FUNCTION_BLOCK "FB_UDP_Pasarela"
{ S7_Optimized_Access := 'TRUE' }
VERSION : 0.1
// PLC_Camara: 279 bloques (un Serialize por miembro de DB o tag). Generado por generar.py
   VAR_INPUT
      Deshabilitar : Bool := FALSE;
      Periodo : Time := T#100ms;
      Ip_pasarela : Array[1..4] of Byte := [172, 21, 0, 200];
      Puerto : UInt := 5000;
   END_VAR
   VAR_OUTPUT
      Conectado : Bool;
      Enviados : UDInt;
      Fallidos : UDInt;
      Bloques_omitidos : Int;
      Estado_tusend : Word;
      Estado_tcon : Word;
      Ultimo_error_tcon : Word;
      Errores_tcon : UDInt;
      Intentos_tcon : UDInt;
      Conexiones_ok : UDInt;
   END_VAR
   VAR
      Etapa : Int;
      Secuencia : UDInt;
      Marca_tiempo : LInt;
      Lanza_conexion : Bool;
      Flanco_conexion : R_TRIG;
      Lanza_envio : Bool;
      Conexion : TCON_IP_v4;
      Destino : TADDR_Param;
      Cliente_con : TCON;
      Cliente_envio : TUSEND;
      Espera_conexion : TON_TIME;
      Espera_periodo : TON_TIME;
      Espera_envio : TON_TIME;
      Datagrama : Array[0..1499] of Byte;
      Foto : Array[0..3384] of Byte;
      Total : DInt;
      Cursor : DInt;
      Bytes_trozo : DInt;
      Bloques_trozo : UInt;
      Bloques_escritos : Int;
      Copia_1 : Array[0..107] of Byte;
      Copia_2 : Bool;
      Copia_3 : Bool;
      Copia_4 : Bool;
      Copia_5 : Bool;
      Copia_6 : Bool;
      Copia_7 : Bool;
      Copia_8 : Bool;
      Copia_9 : Bool;
      Copia_10 : UDInt;
      Copia_11 : UDInt;
      Copia_12 : Bool;
      Copia_13 : Array[0..107] of Byte;
      Copia_14 : UDInt;
      Copia_15 : UDInt;
      Copia_16 : DWord;
      Copia_17 : DWord;
      Copia_18 : DWord;
      Copia_19 : DWord;
      Copia_20 : DWord;
      Copia_21 : DWord;
      Copia_22 : DWord;
      Copia_23 : DWord;
      Copia_24 : DWord;
      Copia_25 : DWord;
      Copia_26 : DWord;
      Copia_27 : DWord;
      Copia_28 : DWord;
      Copia_29 : DWord;
      Copia_30 : DWord;
      Copia_31 : DWord;
      Copia_32 : DWord;
      Copia_33 : DWord;
      Copia_34 : DWord;
      Copia_35 : DWord;
      Copia_36 : DWord;
      Copia_37 : DWord;
      Copia_38 : DWord;
      Copia_39 : DWord;
      Copia_40 : DWord;
      Copia_41 : DWord;
      Copia_42 : DWord;
      Copia_43 : DWord;
      Copia_44 : DWord;
      Copia_45 : DWord;
      Copia_46 : DWord;
      Copia_47 : DWord;
      Copia_48 : Bool;
      Copia_49 : DInt;
      Copia_50 : DInt;
      Copia_51 : Time;
      Copia_52 : "UDT_Entradas_Basico";
      Copia_53 : "UDT_Entradas_RFID";
      Copia_54 : "UDT_Entradas_Stopper";
      Copia_55 : Word;
      Copia_56 : Word;
      Copia_57 : Bool;
      Copia_58 : Bool;
      Copia_59 : Bool;
      Copia_60 : Bool;
      Copia_61 : Bool;
      Copia_62 : DWord;
      Copia_63 : DWord;
      Copia_64 : DWord;
      Copia_65 : DWord;
      Copia_66 : DWord;
      Copia_67 : DWord;
      Copia_68 : DWord;
      Copia_69 : DWord;
      Copia_70 : USInt;
      Copia_71 : UInt;
      Copia_72 : Bool;
      Copia_73 : DInt;
      Copia_74 : Bool;
      Copia_75 : Bool;
      Copia_76 : Bool;
      Copia_77 : UDInt;
      Copia_78 : UDInt;
      Copia_79 : DInt;
      Copia_80 : Int;
      Copia_81 : Bool;
      Copia_82 : Bool;
      Copia_83 : Bool;
      Copia_84 : Bool;
      Copia_85 : Bool;
      Copia_86 : Bool;
      Copia_87 : "UDT_Estado";
      Copia_88 : Bool;
      Copia_89 : Bool;
      Copia_90 : Bool;
      Copia_91 : Bool;
      Copia_92 : Bool;
      Copia_93 : Bool;
      Copia_94 : Bool;
      Copia_95 : Bool;
      Copia_96 : Bool;
      Copia_97 : Bool;
      Copia_98 : Int;
      Copia_99 : Int;
      Copia_100 : Int;
      Copia_101 : Bool;
      Copia_102 : Bool;
      Copia_103 : Bool;
      Copia_104 : Bool;
      Copia_105 : Bool;
      Copia_106 : Bool;
      Copia_107 : Bool;
      Copia_108 : Bool;
      Copia_109 : Bool;
      Copia_110 : Bool;
      Copia_111 : Bool;
      Copia_112 : Bool;
      Copia_113 : Bool;
      Copia_114 : Bool;
      Copia_115 : Bool;
      Copia_116 : Bool;
      Copia_117 : DInt;
      Copia_118 : DInt;
      Copia_119 : Bool;
      Copia_120 : Int;
      Copia_121 : Bool;
      Copia_122 : Bool;
      Copia_123 : Bool;
      Copia_124 : Bool;
      Copia_125 : Int;
      Copia_126 : Bool;
      Copia_127 : Bool;
      Copia_128 : Bool;
      Copia_129 : Bool;
      Copia_130 : Time;
      Copia_131 : Time;
      Copia_132 : Bool;
      Copia_133 : Bool;
      Copia_134 : Time;
      Copia_135 : Time;
      Copia_136 : Bool;
      Copia_137 : Bool;
      Copia_138 : Time;
      Copia_139 : Time;
      Copia_140 : Bool;
      Copia_141 : Bool;
      Copia_142 : Time;
      Copia_143 : Time;
      Copia_144 : Bool;
      Copia_145 : Bool;
      Copia_146 : Bool;
      Copia_147 : Bool;
      Copia_148 : Bool;
      Copia_149 : Bool;
      Copia_150 : Bool;
      Copia_151 : Bool;
      Copia_152 : Bool;
      Copia_153 : Bool;
      Copia_154 : Bool;
      Copia_155 : Bool;
      Copia_156 : Bool;
      Copia_157 : Bool;
      Copia_158 : Byte;
      Copia_159 : Word;
      Copia_160 : Array[0..27] of Byte;
      Copia_161 : Word;
      Copia_162 : Word;
      Copia_163 : DWord;
      Copia_164 : DWord;
      Copia_165 : DWord;
      Copia_166 : DWord;
      Copia_167 : DWord;
      Copia_168 : DWord;
      Copia_169 : DWord;
      Copia_170 : DWord;
      Copia_171 : Bool;
      Copia_172 : Bool;
      Copia_173 : Time;
      Copia_174 : Time;
      Copia_175 : Int;
      Copia_176 : Int;
      Copia_177 : Array[0..3] of DWord;
      Copia_178 : Array[0..3] of DWord;
      Copia_179 : Array[0..3] of Bool;
      Copia_180 : Array[0..3] of Bool;
      Copia_181 : Word;
      Copia_182 : Word;
      Copia_183 : Bool;
      Copia_184 : Bool;
      Copia_185 : Bool;
      Copia_186 : Bool;
      Copia_187 : Bool;
      Copia_188 : Bool;
      Copia_189 : Array[0..107] of Byte;
      Copia_190 : UDInt;
      Copia_191 : UInt;
      Copia_192 : Bool;
      Copia_193 : DTL;
      Copia_194 : Int;
      Copia_195 : DInt;
      Copia_196 : DInt;
      Copia_197 : DInt;
      Copia_198 : DInt;
      Copia_199 : DInt;
      Copia_200 : DInt;
      Copia_201 : DInt;
      Copia_202 : Bool;
      Copia_203 : Bool;
      Copia_204 : Int;
      Copia_205 : Int;
      Copia_206 : UDInt;
      Copia_207 : UInt;
      Copia_208 : UDInt;
      Copia_209 : Bool;
      Copia_210 : Bool;
      Copia_211 : Bool;
      Copia_212 : Time;
      Copia_213 : Time;
      Copia_214 : Bool;
      Copia_215 : Bool;
      Copia_216 : Bool;
      Copia_217 : "UDT_PROFINETSTATUS";
      Copia_218 : "UDT_CAMARA_IN";
      Copia_219 : Bool;
      Copia_220 : Bool;
      Copia_221 : Bool;
      Copia_222 : Bool;
      Copia_223 : Bool;
      Copia_224 : "UDT_PROFINETCTRL";
      Copia_225 : "UDT_CAMARA_OUT";
      Copia_226 : Int;
      Copia_227 : Byte;
      Copia_228 : Bool;
      Copia_229 : Bool;
      Copia_230 : Bool;
      Copia_231 : Bool;
      Copia_232 : Bool;
      Copia_233 : Bool;
      Copia_234 : Bool;
      Copia_235 : Bool;
      Copia_236 : Bool;
      Copia_237 : Bool;
      Copia_238 : Bool;
      Copia_239 : Bool;
      Copia_240 : Time;
      Copia_241 : Time;
      Copia_242 : Bool;
      Copia_243 : Bool;
      Copia_244 : Time;
      Copia_245 : Time;
      Copia_246 : Bool;
      Copia_247 : Bool;
      Copia_248 : Time;
      Copia_249 : Time;
      Copia_250 : Bool;
      Copia_251 : Bool;
      Copia_252 : Time;
      Copia_253 : Time;
      Copia_254 : Bool;
      Copia_255 : Bool;
      Copia_256 : Time;
      Copia_257 : Time;
      Copia_258 : Bool;
      Copia_259 : Bool;
      Copia_260 : Time;
      Copia_261 : Time;
      Copia_262 : UDT_PROFINETCTRL;
      Copia_263 : UDT_PROFINETSTATUS;
      Copia_264 : Byte;
      Copia_265 : Bool;
      Copia_266 : Bool;
      Copia_267 : Bool;
      Copia_268 : Bool;
      Copia_269 : Bool;
      Copia_270 : Bool;
      Copia_271 : Bool;
      Copia_272 : Bool;
      Copia_273 : UDT_CAMARA_IN;
      Copia_274 : UDT_Entradas_Basico;
      Copia_275 : UDT_Entradas_Stopper;
      Copia_276 : UDT_Salidas_Basico;
      Copia_277 : UDT_CAMARA_OUT;
      Copia_278 : UDT_Entradas_RFID;
      Copia_279 : UDT_Salidas_RFID;
   END_VAR
   VAR_TEMP
      periodo_uso : Time;
      puerto_uso : UInt;
      i : Int;
      w : Word;
      d : DWord;
      l : LWord;
      reloj : DTL;
      anio : LInt;
      mes : LInt;
      dia : LInt;
      era : LInt;
      ano_era : LInt;
      dia_ano : LInt;
      dias : LInt;
      resultado : Int;
      longitud : DInt;
      lon_bloque : DInt;
   END_VAR
   VAR CONSTANT
      ID_PLC : USInt := 1;
      N_BLOQUES : Int := 279;
      MAX_PAYLOAD : DInt := 1380;
   END_VAR

BEGIN
// parametros: un valor a cero (DB sin valores iniciales) se sustituye por el de fabrica
#periodo_uso := #Periodo;
IF #periodo_uso <= T#0ms THEN #periodo_uso := T#100ms; END_IF;
#puerto_uso := #Puerto;
IF #puerto_uso = 0 THEN #puerto_uso := 5000; END_IF;

// conexion UDP: un TCON hasta que acabe bien, reintento cada segundo
#Conexion.InterfaceId := "Local~Interfaz_PROFINET_1";
#Conexion.ID := 16#0001;
#Conexion.ConnectionType := 16#13;
#Conexion.ActiveEstablished := FALSE;
#Conexion.RemoteAddress.ADDR := #Ip_pasarela;
#Conexion.RemotePort := #puerto_uso;
#Conexion.LocalPort := #puerto_uso;
FOR #i := 1 TO 4 DO
   #Destino.REM_IP_ADDR[#i] := #Ip_pasarela[#i];
END_FOR;
#Destino.REM_PORT_NR := #puerto_uso;
#Destino.RESERVED := 0;

#Espera_conexion(IN := NOT #Deshabilitar AND NOT #Conectado AND NOT #Cliente_con.BUSY, PT := T#1s);
#Lanza_conexion := #Espera_conexion.Q;
#Cliente_con(REQ := #Lanza_conexion, ID := #Conexion.ID, CONNECT := #Conexion, STATUS => #Estado_tcon);
#Flanco_conexion(CLK := #Lanza_conexion);
IF #Flanco_conexion.Q THEN #Intentos_tcon := #Intentos_tcon + 1; END_IF;
IF #Cliente_con.ERROR THEN
   #Ultimo_error_tcon := #Estado_tcon;
   #Errores_tcon := #Errores_tcon + 1;
END_IF;
IF #Cliente_con.DONE THEN
   IF NOT #Conectado THEN #Conexiones_ok := #Conexiones_ok + 1; END_IF;
   #Conectado := TRUE;
   IF #Etapa = 0 THEN #Etapa := 1; END_IF;
END_IF;
IF #Deshabilitar THEN
   #Conectado := FALSE;
   #Etapa := 0;
END_IF;

// foto de todos los miembros y marca de tiempo UTC (ms desde 1970) cada periodo
#Espera_periodo(IN := #Conectado AND #Etapa = 1, PT := #periodo_uso);
IF #Espera_periodo.Q THEN
   #resultado := RD_SYS_T(OUT => #reloj);
   #anio := UINT_TO_LINT(#reloj.YEAR);
   #mes := USINT_TO_LINT(#reloj.MONTH);
   #dia := USINT_TO_LINT(#reloj.DAY);
   IF #mes <= 2 THEN #anio := #anio - 1; END_IF;
   #era := #anio / 400;
   #ano_era := #anio - #era * 400;
   #dia_ano := (153 * ((#mes + 9) MOD 12) + 2) / 5 + #dia - 1;
   #dias := #era * 146097 + #ano_era * 365 + #ano_era / 4 - #ano_era / 100 + #dia_ano - 719468;
   #Marca_tiempo := ((#dias * 86400 + USINT_TO_LINT(#reloj.HOUR) * 3600 + USINT_TO_LINT(#reloj.MINUTE) * 60
                      + USINT_TO_LINT(#reloj.SECOND)) * 1000) + UDINT_TO_LINT(#reloj.NANOSECOND) / 1000000;
   #Total := 0;
   #Bloques_escritos := 0;
   #Copia_1 := "DB_Estacion".Imagen_palet;
   #Resultado := "FC_UDP_Bloque"(Id := 1, Origen := #Copia_1, Inicio := #Total, Foto := #Foto, Escritos := #Bloques_escritos, Final => #Total);
   #Copia_2 := "DB_Estacion".App_inicio;
   #Resultado := "FC_UDP_Bloque"(Id := 2, Origen := #Copia_2, Inicio := #Total, Foto := #Foto, Escritos := #Bloques_escritos, Final => #Total);
   #Copia_3 := "DB_Estacion".App_en_reposo;
   #Resultado := "FC_UDP_Bloque"(Id := 3, Origen := #Copia_3, Inicio := #Total, Foto := #Foto, Escritos := #Bloques_escritos, Final => #Total);
   #Copia_4 := "DB_Estacion".App_terminada;
   #Resultado := "FC_UDP_Bloque"(Id := 4, Origen := #Copia_4, Inicio := #Total, Foto := #Foto, Escritos := #Bloques_escritos, Final => #Total);
   #Copia_5 := "DB_Estacion".App_alarma;
   #Resultado := "FC_UDP_Bloque"(Id := 5, Origen := #Copia_5, Inicio := #Total, Foto := #Foto, Escritos := #Bloques_escritos, Final => #Total);
   #Copia_6 := "DB_Estacion".App_rearme_requerido;
   #Resultado := "FC_UDP_Bloque"(Id := 6, Origen := #Copia_6, Inicio := #Total, Foto := #Foto, Escritos := #Bloques_escritos, Final => #Total);
   #Copia_7 := "DB_Estacion".Inhibir_cinta;
   #Resultado := "FC_UDP_Bloque"(Id := 7, Origen := #Copia_7, Inicio := #Total, Foto := #Foto, Escritos := #Bloques_escritos, Final => #Total);
   #Copia_8 := "DB_Estacion".Emergencia;
   #Resultado := "FC_UDP_Bloque"(Id := 8, Origen := #Copia_8, Inicio := #Total, Foto := #Foto, Escritos := #Bloques_escritos, Final => #Total);
   #Copia_9 := "DB_Estacion".Rearme;
   #Resultado := "FC_UDP_Bloque"(Id := 9, Origen := #Copia_9, Inicio := #Total, Foto := #Foto, Escritos := #Bloques_escritos, Final => #Total);
   #Copia_10 := "DB_Estacion".Hora_actual;
   #Resultado := "FC_UDP_Bloque"(Id := 10, Origen := #Copia_10, Inicio := #Total, Foto := #Foto, Escritos := #Bloques_escritos, Final => #Total);
   #Copia_11 := "DB_Estacion".Hora_inicio_app;
   #Resultado := "FC_UDP_Bloque"(Id := 11, Origen := #Copia_11, Inicio := #Total, Foto := #Foto, Escritos := #Bloques_escritos, Final => #Total);
   #Copia_12 := "DB_Estacion".Registro_nuevo;
   #Resultado := "FC_UDP_Bloque"(Id := 12, Origen := #Copia_12, Inicio := #Total, Foto := #Foto, Escritos := #Bloques_escritos, Final => #Total);
   #Copia_13 := "DB_Estacion".Registro_palet;
   #Resultado := "FC_UDP_Bloque"(Id := 13, Origen := #Copia_13, Inicio := #Total, Foto := #Foto, Escritos := #Bloques_escritos, Final => #Total);
   #Copia_14 := "DB_Estacion".Out_hora_inicio;
   #Resultado := "FC_UDP_Bloque"(Id := 14, Origen := #Copia_14, Inicio := #Total, Foto := #Foto, Escritos := #Bloques_escritos, Final => #Total);
   #Copia_15 := "DB_Estacion".Out_hora_fin;
   #Resultado := "FC_UDP_Bloque"(Id := 15, Origen := #Copia_15, Inicio := #Total, Foto := #Foto, Escritos := #Bloques_escritos, Final => #Total);
   #Copia_16 := "DB_Estacion".MASCARA_LECTURA_OUT;
   #Resultado := "FC_UDP_Bloque"(Id := 16, Origen := #Copia_16, Inicio := #Total, Foto := #Foto, Escritos := #Bloques_escritos, Final => #Total);
   #Copia_17 := "DB_Estacion".MASCARA_LECTURA_OUT_1;
   #Resultado := "FC_UDP_Bloque"(Id := 17, Origen := #Copia_17, Inicio := #Total, Foto := #Foto, Escritos := #Bloques_escritos, Final => #Total);
   #Copia_18 := "DB_Estacion".MASCARA_LECTURA_OUT_2;
   #Resultado := "FC_UDP_Bloque"(Id := 18, Origen := #Copia_18, Inicio := #Total, Foto := #Foto, Escritos := #Bloques_escritos, Final => #Total);
   #Copia_19 := "DB_Estacion".MASCARA_LECTURA_OUT_3;
   #Resultado := "FC_UDP_Bloque"(Id := 19, Origen := #Copia_19, Inicio := #Total, Foto := #Foto, Escritos := #Bloques_escritos, Final => #Total);
   #Copia_20 := "DB_Estacion".MASCARA_ESCRITURA_OUT;
   #Resultado := "FC_UDP_Bloque"(Id := 20, Origen := #Copia_20, Inicio := #Total, Foto := #Foto, Escritos := #Bloques_escritos, Final => #Total);
   #Copia_21 := "DB_Estacion".MASCARA_ESCRITURA_OUT_1;
   #Resultado := "FC_UDP_Bloque"(Id := 21, Origen := #Copia_21, Inicio := #Total, Foto := #Foto, Escritos := #Bloques_escritos, Final => #Total);
   #Copia_22 := "DB_Estacion".MASCARA_ESCRITURA_OUT_2;
   #Resultado := "FC_UDP_Bloque"(Id := 22, Origen := #Copia_22, Inicio := #Total, Foto := #Foto, Escritos := #Bloques_escritos, Final => #Total);
   #Copia_23 := "DB_Estacion".MASCARA_ESCRITURA_OUT_3;
   #Resultado := "FC_UDP_Bloque"(Id := 23, Origen := #Copia_23, Inicio := #Total, Foto := #Foto, Escritos := #Bloques_escritos, Final => #Total);
   #Copia_24 := "DB_Estacion".MASCARA_LECTURA_PRENSA;
   #Resultado := "FC_UDP_Bloque"(Id := 24, Origen := #Copia_24, Inicio := #Total, Foto := #Foto, Escritos := #Bloques_escritos, Final => #Total);
   #Copia_25 := "DB_Estacion".MASCARA_LECTURA_PRENSA_1;
   #Resultado := "FC_UDP_Bloque"(Id := 25, Origen := #Copia_25, Inicio := #Total, Foto := #Foto, Escritos := #Bloques_escritos, Final => #Total);
   #Copia_26 := "DB_Estacion".MASCARA_LECTURA_PRENSA_2;
   #Resultado := "FC_UDP_Bloque"(Id := 26, Origen := #Copia_26, Inicio := #Total, Foto := #Foto, Escritos := #Bloques_escritos, Final => #Total);
   #Copia_27 := "DB_Estacion".MASCARA_LECTURA_PRENSA_3;
   #Resultado := "FC_UDP_Bloque"(Id := 27, Origen := #Copia_27, Inicio := #Total, Foto := #Foto, Escritos := #Bloques_escritos, Final => #Total);
   #Copia_28 := "DB_Estacion".MASCARA_ESCRITURA_PRENSA;
   #Resultado := "FC_UDP_Bloque"(Id := 28, Origen := #Copia_28, Inicio := #Total, Foto := #Foto, Escritos := #Bloques_escritos, Final => #Total);
   #Copia_29 := "DB_Estacion".MASCARA_ESCRITURA_PRENSA_1;
   #Resultado := "FC_UDP_Bloque"(Id := 29, Origen := #Copia_29, Inicio := #Total, Foto := #Foto, Escritos := #Bloques_escritos, Final => #Total);
   #Copia_30 := "DB_Estacion".MASCARA_ESCRITURA_PRENSA_2;
   #Resultado := "FC_UDP_Bloque"(Id := 30, Origen := #Copia_30, Inicio := #Total, Foto := #Foto, Escritos := #Bloques_escritos, Final => #Total);
   #Copia_31 := "DB_Estacion".MASCARA_ESCRITURA_PRENSA_3;
   #Resultado := "FC_UDP_Bloque"(Id := 31, Origen := #Copia_31, Inicio := #Total, Foto := #Foto, Escritos := #Bloques_escritos, Final => #Total);
   #Copia_32 := "DB_Estacion".MASCARA_LECTURA_CAM;
   #Resultado := "FC_UDP_Bloque"(Id := 32, Origen := #Copia_32, Inicio := #Total, Foto := #Foto, Escritos := #Bloques_escritos, Final => #Total);
   #Copia_33 := "DB_Estacion".MASCARA_LECTURA_CAM_1;
   #Resultado := "FC_UDP_Bloque"(Id := 33, Origen := #Copia_33, Inicio := #Total, Foto := #Foto, Escritos := #Bloques_escritos, Final => #Total);
   #Copia_34 := "DB_Estacion".MASCARA_LECTURA_CAM_2;
   #Resultado := "FC_UDP_Bloque"(Id := 34, Origen := #Copia_34, Inicio := #Total, Foto := #Foto, Escritos := #Bloques_escritos, Final => #Total);
   #Copia_35 := "DB_Estacion".MASCARA_LECTURA_CAM_3;
   #Resultado := "FC_UDP_Bloque"(Id := 35, Origen := #Copia_35, Inicio := #Total, Foto := #Foto, Escritos := #Bloques_escritos, Final => #Total);
   #Copia_36 := "DB_Estacion".MASCARA_ESCRITURA_CAM;
   #Resultado := "FC_UDP_Bloque"(Id := 36, Origen := #Copia_36, Inicio := #Total, Foto := #Foto, Escritos := #Bloques_escritos, Final => #Total);
   #Copia_37 := "DB_Estacion".MASCARA_ESCRITURA_CAM_1;
   #Resultado := "FC_UDP_Bloque"(Id := 37, Origen := #Copia_37, Inicio := #Total, Foto := #Foto, Escritos := #Bloques_escritos, Final => #Total);
   #Copia_38 := "DB_Estacion".MASCARA_ESCRITURA_CAM_2;
   #Resultado := "FC_UDP_Bloque"(Id := 38, Origen := #Copia_38, Inicio := #Total, Foto := #Foto, Escritos := #Bloques_escritos, Final => #Total);
   #Copia_39 := "DB_Estacion".MASCARA_ESCRITURA_CAM_3;
   #Resultado := "FC_UDP_Bloque"(Id := 39, Origen := #Copia_39, Inicio := #Total, Foto := #Foto, Escritos := #Bloques_escritos, Final => #Total);
   #Copia_40 := "DB_Estacion".MASCARA_LECTURA_BACK;
   #Resultado := "FC_UDP_Bloque"(Id := 40, Origen := #Copia_40, Inicio := #Total, Foto := #Foto, Escritos := #Bloques_escritos, Final => #Total);
   #Copia_41 := "DB_Estacion".MASCARA_LECTURA_BACK_1;
   #Resultado := "FC_UDP_Bloque"(Id := 41, Origen := #Copia_41, Inicio := #Total, Foto := #Foto, Escritos := #Bloques_escritos, Final => #Total);
   #Copia_42 := "DB_Estacion".MASCARA_LECTURA_BACK_2;
   #Resultado := "FC_UDP_Bloque"(Id := 42, Origen := #Copia_42, Inicio := #Total, Foto := #Foto, Escritos := #Bloques_escritos, Final => #Total);
   #Copia_43 := "DB_Estacion".MASCARA_LECTURA_BACK_3;
   #Resultado := "FC_UDP_Bloque"(Id := 43, Origen := #Copia_43, Inicio := #Total, Foto := #Foto, Escritos := #Bloques_escritos, Final => #Total);
   #Copia_44 := "DB_Estacion".MASCARA_ESCRITURA_BACK;
   #Resultado := "FC_UDP_Bloque"(Id := 44, Origen := #Copia_44, Inicio := #Total, Foto := #Foto, Escritos := #Bloques_escritos, Final => #Total);
   #Copia_45 := "DB_Estacion".MASCARA_ESCRITURA_BACK_1;
   #Resultado := "FC_UDP_Bloque"(Id := 45, Origen := #Copia_45, Inicio := #Total, Foto := #Foto, Escritos := #Bloques_escritos, Final => #Total);
   #Copia_46 := "DB_Estacion".MASCARA_ESCRITURA_BACK_2;
   #Resultado := "FC_UDP_Bloque"(Id := 46, Origen := #Copia_46, Inicio := #Total, Foto := #Foto, Escritos := #Bloques_escritos, Final => #Total);
   #Copia_47 := "DB_Estacion".MASCARA_ESCRITURA_BACK_3;
   #Resultado := "FC_UDP_Bloque"(Id := 47, Origen := #Copia_47, Inicio := #Total, Foto := #Foto, Escritos := #Bloques_escritos, Final => #Total);
   #Copia_48 := "DB_Estacion".Parada_fina;
   #Resultado := "FC_UDP_Bloque"(Id := 48, Origen := #Copia_48, Inicio := #Total, Foto := #Foto, Escritos := #Bloques_escritos, Final => #Total);
   #Copia_49 := "DB_Estacion".Encoder_cuentas;
   #Resultado := "FC_UDP_Bloque"(Id := 49, Origen := #Copia_49, Inicio := #Total, Foto := #Foto, Escritos := #Bloques_escritos, Final => #Total);
   #Copia_50 := "DB_Estacion".Distancia_parada_fina_cuentas;
   #Resultado := "FC_UDP_Bloque"(Id := 50, Origen := #Copia_50, Inicio := #Total, Foto := #Foto, Escritos := #Bloques_escritos, Final => #Total);
   #Copia_51 := "DB_Estacion".Tiempo_bajada_cilindro;
   #Resultado := "FC_UDP_Bloque"(Id := 51, Origen := #Copia_51, Inicio := #Total, Foto := #Foto, Escritos := #Bloques_escritos, Final => #Total);
   #Copia_52 := "Est_DB_Gestor".InBasico;
   #Resultado := "FC_UDP_Bloque"(Id := 52, Origen := #Copia_52, Inicio := #Total, Foto := #Foto, Escritos := #Bloques_escritos, Final => #Total);
   #Copia_53 := "Est_DB_Gestor".InRFID;
   #Resultado := "FC_UDP_Bloque"(Id := 53, Origen := #Copia_53, Inicio := #Total, Foto := #Foto, Escritos := #Bloques_escritos, Final => #Total);
   #Copia_54 := "Est_DB_Gestor".InStopper;
   #Resultado := "FC_UDP_Bloque"(Id := 54, Origen := #Copia_54, Inicio := #Total, Foto := #Foto, Escritos := #Bloques_escritos, Final => #Total);
   #Copia_55 := "Est_DB_Gestor".Direccion_lectura;
   #Resultado := "FC_UDP_Bloque"(Id := 55, Origen := #Copia_55, Inicio := #Total, Foto := #Foto, Escritos := #Bloques_escritos, Final => #Total);
   #Copia_56 := "Est_DB_Gestor".Direccion_escritura;
   #Resultado := "FC_UDP_Bloque"(Id := 56, Origen := #Copia_56, Inicio := #Total, Foto := #Foto, Escritos := #Bloques_escritos, Final => #Total);
   #Copia_57 := "Est_DB_Gestor".App_en_reposo;
   #Resultado := "FC_UDP_Bloque"(Id := 57, Origen := #Copia_57, Inicio := #Total, Foto := #Foto, Escritos := #Bloques_escritos, Final => #Total);
   #Copia_58 := "Est_DB_Gestor".App_terminada;
   #Resultado := "FC_UDP_Bloque"(Id := 58, Origen := #Copia_58, Inicio := #Total, Foto := #Foto, Escritos := #Bloques_escritos, Final => #Total);
   #Copia_59 := "Est_DB_Gestor".App_alarma;
   #Resultado := "FC_UDP_Bloque"(Id := 59, Origen := #Copia_59, Inicio := #Total, Foto := #Foto, Escritos := #Bloques_escritos, Final => #Total);
   #Copia_60 := "Est_DB_Gestor".App_rearme_requerido;
   #Resultado := "FC_UDP_Bloque"(Id := 60, Origen := #Copia_60, Inicio := #Total, Foto := #Foto, Escritos := #Bloques_escritos, Final => #Total);
   #Copia_61 := "Est_DB_Gestor".Inhibir_cinta;
   #Resultado := "FC_UDP_Bloque"(Id := 61, Origen := #Copia_61, Inicio := #Total, Foto := #Foto, Escritos := #Bloques_escritos, Final => #Total);
   #Copia_62 := "Est_DB_Gestor".Mascara_lectura;
   #Resultado := "FC_UDP_Bloque"(Id := 62, Origen := #Copia_62, Inicio := #Total, Foto := #Foto, Escritos := #Bloques_escritos, Final => #Total);
   #Copia_63 := "Est_DB_Gestor".Mascara_escritura;
   #Resultado := "FC_UDP_Bloque"(Id := 63, Origen := #Copia_63, Inicio := #Total, Foto := #Foto, Escritos := #Bloques_escritos, Final => #Total);
   #Copia_64 := "Est_DB_Gestor".Mascara_lectura_1;
   #Resultado := "FC_UDP_Bloque"(Id := 64, Origen := #Copia_64, Inicio := #Total, Foto := #Foto, Escritos := #Bloques_escritos, Final => #Total);
   #Copia_65 := "Est_DB_Gestor".Mascara_lectura_2;
   #Resultado := "FC_UDP_Bloque"(Id := 65, Origen := #Copia_65, Inicio := #Total, Foto := #Foto, Escritos := #Bloques_escritos, Final => #Total);
   #Copia_66 := "Est_DB_Gestor".Mascara_lectura_3;
   #Resultado := "FC_UDP_Bloque"(Id := 66, Origen := #Copia_66, Inicio := #Total, Foto := #Foto, Escritos := #Bloques_escritos, Final => #Total);
   #Copia_67 := "Est_DB_Gestor".Mascara_escritura_1;
   #Resultado := "FC_UDP_Bloque"(Id := 67, Origen := #Copia_67, Inicio := #Total, Foto := #Foto, Escritos := #Bloques_escritos, Final => #Total);
   #Copia_68 := "Est_DB_Gestor".Mascara_escritura_2;
   #Resultado := "FC_UDP_Bloque"(Id := 68, Origen := #Copia_68, Inicio := #Total, Foto := #Foto, Escritos := #Bloques_escritos, Final => #Total);
   #Copia_69 := "Est_DB_Gestor".Mascara_escritura_3;
   #Resultado := "FC_UDP_Bloque"(Id := 69, Origen := #Copia_69, Inicio := #Total, Foto := #Foto, Escritos := #Bloques_escritos, Final => #Total);
   #Copia_70 := "Est_DB_Gestor".Id_estacion;
   #Resultado := "FC_UDP_Bloque"(Id := 70, Origen := #Copia_70, Inicio := #Total, Foto := #Foto, Escritos := #Bloques_escritos, Final => #Total);
   #Copia_71 := "Est_DB_Gestor".Lote;
   #Resultado := "FC_UDP_Bloque"(Id := 71, Origen := #Copia_71, Inicio := #Total, Foto := #Foto, Escritos := #Bloques_escritos, Final => #Total);
   #Copia_72 := "Est_DB_Gestor".Parada_fina;
   #Resultado := "FC_UDP_Bloque"(Id := 72, Origen := #Copia_72, Inicio := #Total, Foto := #Foto, Escritos := #Bloques_escritos, Final => #Total);
   #Copia_73 := "Est_DB_Gestor".Distancia_parada_fina_cuentas;
   #Resultado := "FC_UDP_Bloque"(Id := 73, Origen := #Copia_73, Inicio := #Total, Foto := #Foto, Escritos := #Bloques_escritos, Final => #Total);
   #Copia_74 := "Est_DB_Gestor".App_inicio;
   #Resultado := "FC_UDP_Bloque"(Id := 74, Origen := #Copia_74, Inicio := #Total, Foto := #Foto, Escritos := #Bloques_escritos, Final => #Total);
   #Copia_75 := "Est_DB_Gestor".Emergencia;
   #Resultado := "FC_UDP_Bloque"(Id := 75, Origen := #Copia_75, Inicio := #Total, Foto := #Foto, Escritos := #Bloques_escritos, Final => #Total);
   #Copia_76 := "Est_DB_Gestor".Rearme;
   #Resultado := "FC_UDP_Bloque"(Id := 76, Origen := #Copia_76, Inicio := #Total, Foto := #Foto, Escritos := #Bloques_escritos, Final => #Total);
   #Copia_77 := "Est_DB_Gestor".Hora_actual;
   #Resultado := "FC_UDP_Bloque"(Id := 77, Origen := #Copia_77, Inicio := #Total, Foto := #Foto, Escritos := #Bloques_escritos, Final => #Total);
   #Copia_78 := "Est_DB_Gestor".Hora_inicio_app;
   #Resultado := "FC_UDP_Bloque"(Id := 78, Origen := #Copia_78, Inicio := #Total, Foto := #Foto, Escritos := #Bloques_escritos, Final => #Total);
   #Copia_79 := "Est_DB_Gestor".Encoder_cuentas;
   #Resultado := "FC_UDP_Bloque"(Id := 79, Origen := #Copia_79, Inicio := #Total, Foto := #Foto, Escritos := #Bloques_escritos, Final => #Total);
   #Copia_80 := "Est_DB_Gestor".Etapa_gestion;
   #Resultado := "FC_UDP_Bloque"(Id := 80, Origen := #Copia_80, Inicio := #Total, Foto := #Foto, Escritos := #Bloques_escritos, Final => #Total);
   #Copia_81 := "Est_DB_Gestor".Etapa_0;
   #Resultado := "FC_UDP_Bloque"(Id := 81, Origen := #Copia_81, Inicio := #Total, Foto := #Foto, Escritos := #Bloques_escritos, Final => #Total);
   #Copia_82 := "Est_DB_Gestor".Etapa_1;
   #Resultado := "FC_UDP_Bloque"(Id := 82, Origen := #Copia_82, Inicio := #Total, Foto := #Foto, Escritos := #Bloques_escritos, Final => #Total);
   #Copia_83 := "Est_DB_Gestor".Etapa_2;
   #Resultado := "FC_UDP_Bloque"(Id := 83, Origen := #Copia_83, Inicio := #Total, Foto := #Foto, Escritos := #Bloques_escritos, Final => #Total);
   #Copia_84 := "Est_DB_Gestor".Etapa_3;
   #Resultado := "FC_UDP_Bloque"(Id := 84, Origen := #Copia_84, Inicio := #Total, Foto := #Foto, Escritos := #Bloques_escritos, Final => #Total);
   #Copia_85 := "Est_DB_Gestor".Etapa_4;
   #Resultado := "FC_UDP_Bloque"(Id := 85, Origen := #Copia_85, Inicio := #Total, Foto := #Foto, Escritos := #Bloques_escritos, Final => #Total);
   #Copia_86 := "Est_DB_Gestor".Etapa_5;
   #Resultado := "FC_UDP_Bloque"(Id := 86, Origen := #Copia_86, Inicio := #Total, Foto := #Foto, Escritos := #Bloques_escritos, Final => #Total);
   #Copia_87 := "Est_DB_Gestor".Estado_Estacion;
   #Resultado := "FC_UDP_Bloque"(Id := 87, Origen := #Copia_87, Inicio := #Total, Foto := #Foto, Escritos := #Bloques_escritos, Final => #Total);
   #Copia_88 := "Est_DB_Gestor".Flanco_rearme.CLK;
   #Resultado := "FC_UDP_Bloque"(Id := 88, Origen := #Copia_88, Inicio := #Total, Foto := #Foto, Escritos := #Bloques_escritos, Final => #Total);
   #Copia_89 := "Est_DB_Gestor".Flanco_rearme.Q;
   #Resultado := "FC_UDP_Bloque"(Id := 89, Origen := #Copia_89, Inicio := #Total, Foto := #Foto, Escritos := #Bloques_escritos, Final => #Total);
   #Copia_90 := "Est_DB_Gestor".FB2_Modo_Instance.Seta_emergencia;
   #Resultado := "FC_UDP_Bloque"(Id := 90, Origen := #Copia_90, Inicio := #Total, Foto := #Foto, Escritos := #Bloques_escritos, Final => #Total);
   #Copia_91 := "Est_DB_Gestor".FB2_Modo_Instance.Boton_rearme;
   #Resultado := "FC_UDP_Bloque"(Id := 91, Origen := #Copia_91, Inicio := #Total, Foto := #Foto, Escritos := #Bloques_escritos, Final => #Total);
   #Copia_92 := "Est_DB_Gestor".FB2_Modo_Instance.Boton_marcha;
   #Resultado := "FC_UDP_Bloque"(Id := 92, Origen := #Copia_92, Inicio := #Total, Foto := #Foto, Escritos := #Bloques_escritos, Final => #Total);
   #Copia_93 := "Est_DB_Gestor".FB2_Modo_Instance.Boton_paro;
   #Resultado := "FC_UDP_Bloque"(Id := 93, Origen := #Copia_93, Inicio := #Total, Foto := #Foto, Escritos := #Bloques_escritos, Final => #Total);
   #Copia_94 := "Est_DB_Gestor".FB2_Modo_Instance.Selector_automatico;
   #Resultado := "FC_UDP_Bloque"(Id := 94, Origen := #Copia_94, Inicio := #Total, Foto := #Foto, Escritos := #Bloques_escritos, Final => #Total);
   #Copia_95 := "Est_DB_Gestor".FB2_Modo_Instance.Condicion_arranque_auto;
   #Resultado := "FC_UDP_Bloque"(Id := 95, Origen := #Copia_95, Inicio := #Total, Foto := #Foto, Escritos := #Bloques_escritos, Final => #Total);
   #Copia_96 := "Est_DB_Gestor".FB2_Modo_Instance.Condicion_arranque_manual;
   #Resultado := "FC_UDP_Bloque"(Id := 96, Origen := #Copia_96, Inicio := #Total, Foto := #Foto, Escritos := #Bloques_escritos, Final => #Total);
   #Copia_97 := "Est_DB_Gestor".FB2_Modo_Instance.Ciclo_manual_acabado;
   #Resultado := "FC_UDP_Bloque"(Id := 97, Origen := #Copia_97, Inicio := #Total, Foto := #Foto, Escritos := #Bloques_escritos, Final => #Total);
   #Copia_98 := "Est_DB_Gestor".FB2_Modo_Instance.Etapa_emergencia;
   #Resultado := "FC_UDP_Bloque"(Id := 98, Origen := #Copia_98, Inicio := #Total, Foto := #Foto, Escritos := #Bloques_escritos, Final => #Total);
   #Copia_99 := "Est_DB_Gestor".FB2_Modo_Instance.Etapa_modo;
   #Resultado := "FC_UDP_Bloque"(Id := 99, Origen := #Copia_99, Inicio := #Total, Foto := #Foto, Escritos := #Bloques_escritos, Final => #Total);
   #Copia_100 := "Est_DB_Gestor".FB2_Modo_Instance.Etapa_ciclo;
   #Resultado := "FC_UDP_Bloque"(Id := 100, Origen := #Copia_100, Inicio := #Total, Foto := #Foto, Escritos := #Bloques_escritos, Final => #Total);
   #Copia_101 := "Est_DB_Gestor".FB2_Modo_Instance.Flanco_marcha.CLK;
   #Resultado := "FC_UDP_Bloque"(Id := 101, Origen := #Copia_101, Inicio := #Total, Foto := #Foto, Escritos := #Bloques_escritos, Final => #Total);
   #Copia_102 := "Est_DB_Gestor".FB2_Modo_Instance.Flanco_marcha.Q;
   #Resultado := "FC_UDP_Bloque"(Id := 102, Origen := #Copia_102, Inicio := #Total, Foto := #Foto, Escritos := #Bloques_escritos, Final => #Total);
   #Copia_103 := "Est_DB_Gestor".FB2_Modo_Instance.Flanco_rearme.CLK;
   #Resultado := "FC_UDP_Bloque"(Id := 103, Origen := #Copia_103, Inicio := #Total, Foto := #Foto, Escritos := #Bloques_escritos, Final => #Total);
   #Copia_104 := "Est_DB_Gestor".FB2_Modo_Instance.Flanco_rearme.Q;
   #Resultado := "FC_UDP_Bloque"(Id := 104, Origen := #Copia_104, Inicio := #Total, Foto := #Foto, Escritos := #Bloques_escritos, Final => #Total);
   #Copia_105 := "Est_DB_Gestor".FB3_Cinta_Instance.Emergencia;
   #Resultado := "FC_UDP_Bloque"(Id := 105, Origen := #Copia_105, Inicio := #Total, Foto := #Foto, Escritos := #Bloques_escritos, Final => #Total);
   #Copia_106 := "Est_DB_Gestor".FB3_Cinta_Instance.Cinta_habilitada;
   #Resultado := "FC_UDP_Bloque"(Id := 106, Origen := #Copia_106, Inicio := #Total, Foto := #Foto, Escritos := #Bloques_escritos, Final => #Total);
   #Copia_107 := "Est_DB_Gestor".FB3_Cinta_Instance.Orden_evacuar;
   #Resultado := "FC_UDP_Bloque"(Id := 107, Origen := #Copia_107, Inicio := #Total, Foto := #Foto, Escritos := #Bloques_escritos, Final => #Total);
   #Copia_108 := "Est_DB_Gestor".FB3_Cinta_Instance.Sensor_palet_izq;
   #Resultado := "FC_UDP_Bloque"(Id := 108, Origen := #Copia_108, Inicio := #Total, Foto := #Foto, Escritos := #Bloques_escritos, Final => #Total);
   #Copia_109 := "Est_DB_Gestor".FB3_Cinta_Instance.Sensor_palet_dch;
   #Resultado := "FC_UDP_Bloque"(Id := 109, Origen := #Copia_109, Inicio := #Total, Foto := #Foto, Escritos := #Bloques_escritos, Final => #Total);
   #Copia_110 := "Est_DB_Gestor".FB3_Cinta_Instance.Sensor_ind_bien_pos;
   #Resultado := "FC_UDP_Bloque"(Id := 110, Origen := #Copia_110, Inicio := #Total, Foto := #Foto, Escritos := #Bloques_escritos, Final => #Total);
   #Copia_111 := "Est_DB_Gestor".FB3_Cinta_Instance.Sensor_stopper_abajo;
   #Resultado := "FC_UDP_Bloque"(Id := 111, Origen := #Copia_111, Inicio := #Total, Foto := #Foto, Escritos := #Bloques_escritos, Final => #Total);
   #Copia_112 := "Est_DB_Gestor".FB3_Cinta_Instance.Sensor_ind_1;
   #Resultado := "FC_UDP_Bloque"(Id := 112, Origen := #Copia_112, Inicio := #Total, Foto := #Foto, Escritos := #Bloques_escritos, Final => #Total);
   #Copia_113 := "Est_DB_Gestor".FB3_Cinta_Instance.Sensor_ind_2;
   #Resultado := "FC_UDP_Bloque"(Id := 113, Origen := #Copia_113, Inicio := #Total, Foto := #Foto, Escritos := #Bloques_escritos, Final => #Total);
   #Copia_114 := "Est_DB_Gestor".FB3_Cinta_Instance.Sensor_ind_3;
   #Resultado := "FC_UDP_Bloque"(Id := 114, Origen := #Copia_114, Inicio := #Total, Foto := #Foto, Escritos := #Bloques_escritos, Final => #Total);
   #Copia_115 := "Est_DB_Gestor".FB3_Cinta_Instance.Parada_fina;
   #Resultado := "FC_UDP_Bloque"(Id := 115, Origen := #Copia_115, Inicio := #Total, Foto := #Foto, Escritos := #Bloques_escritos, Final => #Total);
   #Copia_116 := "Est_DB_Gestor".FB3_Cinta_Instance.Encoder_A;
   #Resultado := "FC_UDP_Bloque"(Id := 116, Origen := #Copia_116, Inicio := #Total, Foto := #Foto, Escritos := #Bloques_escritos, Final => #Total);
   #Copia_117 := "Est_DB_Gestor".FB3_Cinta_Instance.Distancia_parada_fina_cuentas;
   #Resultado := "FC_UDP_Bloque"(Id := 117, Origen := #Copia_117, Inicio := #Total, Foto := #Foto, Escritos := #Bloques_escritos, Final => #Total);
   #Copia_118 := "Est_DB_Gestor".FB3_Cinta_Instance.Encoder_cuentas;
   #Resultado := "FC_UDP_Bloque"(Id := 118, Origen := #Copia_118, Inicio := #Total, Foto := #Foto, Escritos := #Bloques_escritos, Final => #Total);
   #Copia_119 := "Est_DB_Gestor".FB3_Cinta_Instance.Velocidad_baja;
   #Resultado := "FC_UDP_Bloque"(Id := 119, Origen := #Copia_119, Inicio := #Total, Foto := #Foto, Escritos := #Bloques_escritos, Final => #Total);
   #Copia_120 := "Est_DB_Gestor".FB3_Cinta_Instance.Etapa_cinta;
   #Resultado := "FC_UDP_Bloque"(Id := 120, Origen := #Copia_120, Inicio := #Total, Foto := #Foto, Escritos := #Bloques_escritos, Final => #Total);
   #Copia_121 := "Est_DB_Gestor".FB3_Cinta_Instance.Flanco_subida_sensor_palet_dch.CLK;
   #Resultado := "FC_UDP_Bloque"(Id := 121, Origen := #Copia_121, Inicio := #Total, Foto := #Foto, Escritos := #Bloques_escritos, Final => #Total);
   #Copia_122 := "Est_DB_Gestor".FB3_Cinta_Instance.Flanco_subida_sensor_palet_dch.Q;
   #Resultado := "FC_UDP_Bloque"(Id := 122, Origen := #Copia_122, Inicio := #Total, Foto := #Foto, Escritos := #Bloques_escritos, Final => #Total);
   #Copia_123 := "Est_DB_Gestor".FB3_Cinta_Instance.Flanco_bajada_sensor_palet_dch.CLK;
   #Resultado := "FC_UDP_Bloque"(Id := 123, Origen := #Copia_123, Inicio := #Total, Foto := #Foto, Escritos := #Bloques_escritos, Final => #Total);
   #Copia_124 := "Est_DB_Gestor".FB3_Cinta_Instance.Flanco_bajada_sensor_palet_dch.Q;
   #Resultado := "FC_UDP_Bloque"(Id := 124, Origen := #Copia_124, Inicio := #Total, Foto := #Foto, Escritos := #Bloques_escritos, Final => #Total);
   #Copia_125 := "Est_DB_Gestor".FB3_Cinta_Instance.Palets_en_cinta;
   #Resultado := "FC_UDP_Bloque"(Id := 125, Origen := #Copia_125, Inicio := #Total, Foto := #Foto, Escritos := #Bloques_escritos, Final => #Total);
   #Copia_126 := "Est_DB_Gestor".FB3_Cinta_Instance.Flanco_subida_sensor_palet_izq.CLK;
   #Resultado := "FC_UDP_Bloque"(Id := 126, Origen := #Copia_126, Inicio := #Total, Foto := #Foto, Escritos := #Bloques_escritos, Final => #Total);
   #Copia_127 := "Est_DB_Gestor".FB3_Cinta_Instance.Flanco_subida_sensor_palet_izq.Q;
   #Resultado := "FC_UDP_Bloque"(Id := 127, Origen := #Copia_127, Inicio := #Total, Foto := #Foto, Escritos := #Bloques_escritos, Final => #Total);
   #Copia_128 := "Est_DB_Gestor".FB3_Cinta_Instance.Timer_Stopper_Etapa5.IN;
   #Resultado := "FC_UDP_Bloque"(Id := 128, Origen := #Copia_128, Inicio := #Total, Foto := #Foto, Escritos := #Bloques_escritos, Final => #Total);
   #Copia_129 := "Est_DB_Gestor".FB3_Cinta_Instance.Timer_Stopper_Etapa5.Q;
   #Resultado := "FC_UDP_Bloque"(Id := 129, Origen := #Copia_129, Inicio := #Total, Foto := #Foto, Escritos := #Bloques_escritos, Final => #Total);
   #Copia_130 := "Est_DB_Gestor".FB3_Cinta_Instance.Timer_Stopper_Etapa5.PT;
   #Resultado := "FC_UDP_Bloque"(Id := 130, Origen := #Copia_130, Inicio := #Total, Foto := #Foto, Escritos := #Bloques_escritos, Final => #Total);
   #Copia_131 := "Est_DB_Gestor".FB3_Cinta_Instance.Timer_Stopper_Etapa5.ET;
   #Resultado := "FC_UDP_Bloque"(Id := 131, Origen := #Copia_131, Inicio := #Total, Foto := #Foto, Escritos := #Bloques_escritos, Final => #Total);
   #Copia_132 := "Est_DB_Gestor".FB3_Cinta_Instance.Timer_avance.IN;
   #Resultado := "FC_UDP_Bloque"(Id := 132, Origen := #Copia_132, Inicio := #Total, Foto := #Foto, Escritos := #Bloques_escritos, Final => #Total);
   #Copia_133 := "Est_DB_Gestor".FB3_Cinta_Instance.Timer_avance.Q;
   #Resultado := "FC_UDP_Bloque"(Id := 133, Origen := #Copia_133, Inicio := #Total, Foto := #Foto, Escritos := #Bloques_escritos, Final => #Total);
   #Copia_134 := "Est_DB_Gestor".FB3_Cinta_Instance.Timer_avance.PT;
   #Resultado := "FC_UDP_Bloque"(Id := 134, Origen := #Copia_134, Inicio := #Total, Foto := #Foto, Escritos := #Bloques_escritos, Final => #Total);
   #Copia_135 := "Est_DB_Gestor".FB3_Cinta_Instance.Timer_avance.ET;
   #Resultado := "FC_UDP_Bloque"(Id := 135, Origen := #Copia_135, Inicio := #Total, Foto := #Foto, Escritos := #Bloques_escritos, Final => #Total);
   #Copia_136 := "Est_DB_Gestor".FB3_Cinta_Instance.Timer_salida_extra.IN;
   #Resultado := "FC_UDP_Bloque"(Id := 136, Origen := #Copia_136, Inicio := #Total, Foto := #Foto, Escritos := #Bloques_escritos, Final => #Total);
   #Copia_137 := "Est_DB_Gestor".FB3_Cinta_Instance.Timer_salida_extra.Q;
   #Resultado := "FC_UDP_Bloque"(Id := 137, Origen := #Copia_137, Inicio := #Total, Foto := #Foto, Escritos := #Bloques_escritos, Final => #Total);
   #Copia_138 := "Est_DB_Gestor".FB3_Cinta_Instance.Timer_salida_extra.PT;
   #Resultado := "FC_UDP_Bloque"(Id := 138, Origen := #Copia_138, Inicio := #Total, Foto := #Foto, Escritos := #Bloques_escritos, Final => #Total);
   #Copia_139 := "Est_DB_Gestor".FB3_Cinta_Instance.Timer_salida_extra.ET;
   #Resultado := "FC_UDP_Bloque"(Id := 139, Origen := #Copia_139, Inicio := #Total, Foto := #Foto, Escritos := #Bloques_escritos, Final => #Total);
   #Copia_140 := "Est_DB_Gestor".FB3_Cinta_Instance.Timer_parada_fina.IN;
   #Resultado := "FC_UDP_Bloque"(Id := 140, Origen := #Copia_140, Inicio := #Total, Foto := #Foto, Escritos := #Bloques_escritos, Final => #Total);
   #Copia_141 := "Est_DB_Gestor".FB3_Cinta_Instance.Timer_parada_fina.Q;
   #Resultado := "FC_UDP_Bloque"(Id := 141, Origen := #Copia_141, Inicio := #Total, Foto := #Foto, Escritos := #Bloques_escritos, Final => #Total);
   #Copia_142 := "Est_DB_Gestor".FB3_Cinta_Instance.Timer_parada_fina.PT;
   #Resultado := "FC_UDP_Bloque"(Id := 142, Origen := #Copia_142, Inicio := #Total, Foto := #Foto, Escritos := #Bloques_escritos, Final => #Total);
   #Copia_143 := "Est_DB_Gestor".FB3_Cinta_Instance.Timer_parada_fina.ET;
   #Resultado := "FC_UDP_Bloque"(Id := 143, Origen := #Copia_143, Inicio := #Total, Foto := #Foto, Escritos := #Bloques_escritos, Final => #Total);
   #Copia_144 := "Est_DB_Gestor".FB3_Cinta_Instance.Flanco_encoder_A.CLK;
   #Resultado := "FC_UDP_Bloque"(Id := 144, Origen := #Copia_144, Inicio := #Total, Foto := #Foto, Escritos := #Bloques_escritos, Final => #Total);
   #Copia_145 := "Est_DB_Gestor".FB3_Cinta_Instance.Flanco_encoder_A.Q;
   #Resultado := "FC_UDP_Bloque"(Id := 145, Origen := #Copia_145, Inicio := #Total, Foto := #Foto, Escritos := #Bloques_escritos, Final => #Total);
   #Copia_146 := "Est_DB_Gestor".FB3_Cinta_Instance.Flanco_sensor_ind_bien_pos.CLK;
   #Resultado := "FC_UDP_Bloque"(Id := 146, Origen := #Copia_146, Inicio := #Total, Foto := #Foto, Escritos := #Bloques_escritos, Final => #Total);
   #Copia_147 := "Est_DB_Gestor".FB3_Cinta_Instance.Flanco_sensor_ind_bien_pos.Q;
   #Resultado := "FC_UDP_Bloque"(Id := 147, Origen := #Copia_147, Inicio := #Total, Foto := #Foto, Escritos := #Bloques_escritos, Final => #Total);
   #Copia_148 := "Est_DB_Gestor".FB3_Cinta_Instance.Aviso_lento;
   #Resultado := "FC_UDP_Bloque"(Id := 148, Origen := #Copia_148, Inicio := #Total, Foto := #Foto, Escritos := #Bloques_escritos, Final => #Total);
   #Copia_149 := "Est_DB_Gestor".FB4_RFID_Instance.Emergencia;
   #Resultado := "FC_UDP_Bloque"(Id := 149, Origen := #Copia_149, Inicio := #Total, Foto := #Foto, Escritos := #Bloques_escritos, Final => #Total);
   #Copia_150 := "Est_DB_Gestor".FB4_RFID_Instance.Orden_escribir;
   #Resultado := "FC_UDP_Bloque"(Id := 150, Origen := #Copia_150, Inicio := #Total, Foto := #Foto, Escritos := #Bloques_escritos, Final => #Total);
   #Copia_151 := "Est_DB_Gestor".FB4_RFID_Instance.Orden_leer;
   #Resultado := "FC_UDP_Bloque"(Id := 151, Origen := #Copia_151, Inicio := #Total, Foto := #Foto, Escritos := #Bloques_escritos, Final => #Total);
   #Copia_152 := "Est_DB_Gestor".FB4_RFID_Instance.Tag_datos_escritos;
   #Resultado := "FC_UDP_Bloque"(Id := 152, Origen := #Copia_152, Inicio := #Total, Foto := #Foto, Escritos := #Bloques_escritos, Final => #Total);
   #Copia_153 := "Est_DB_Gestor".FB4_RFID_Instance.Tag_datos_leidos;
   #Resultado := "FC_UDP_Bloque"(Id := 153, Origen := #Copia_153, Inicio := #Total, Foto := #Foto, Escritos := #Bloques_escritos, Final => #Total);
   #Copia_154 := "Est_DB_Gestor".FB4_RFID_Instance.Tag_antena_apagada;
   #Resultado := "FC_UDP_Bloque"(Id := 154, Origen := #Copia_154, Inicio := #Total, Foto := #Foto, Escritos := #Bloques_escritos, Final => #Total);
   #Copia_155 := "Est_DB_Gestor".FB4_RFID_Instance.Tag_detectado;
   #Resultado := "FC_UDP_Bloque"(Id := 155, Origen := #Copia_155, Inicio := #Total, Foto := #Foto, Escritos := #Bloques_escritos, Final => #Total);
   #Copia_156 := "Est_DB_Gestor".FB4_RFID_Instance.Tag_error;
   #Resultado := "FC_UDP_Bloque"(Id := 156, Origen := #Copia_156, Inicio := #Total, Foto := #Foto, Escritos := #Bloques_escritos, Final => #Total);
   #Copia_157 := "Est_DB_Gestor".FB4_RFID_Instance.Tag_proceso_listo;
   #Resultado := "FC_UDP_Bloque"(Id := 157, Origen := #Copia_157, Inicio := #Total, Foto := #Foto, Escritos := #Bloques_escritos, Final => #Total);
   #Copia_158 := "Est_DB_Gestor".FB4_RFID_Instance.Tag_codigo_error;
   #Resultado := "FC_UDP_Bloque"(Id := 158, Origen := #Copia_158, Inicio := #Total, Foto := #Foto, Escritos := #Bloques_escritos, Final => #Total);
   #Copia_159 := "Est_DB_Gestor".FB4_RFID_Instance.Tag_direccion_confirmada;
   #Resultado := "FC_UDP_Bloque"(Id := 159, Origen := #Copia_159, Inicio := #Total, Foto := #Foto, Escritos := #Bloques_escritos, Final => #Total);
   #Copia_160 := "Est_DB_Gestor".FB4_RFID_Instance.Tag_datos_leidos_escritos;
   #Resultado := "FC_UDP_Bloque"(Id := 160, Origen := #Copia_160, Inicio := #Total, Foto := #Foto, Escritos := #Bloques_escritos, Final => #Total);
   #Copia_161 := "Est_DB_Gestor".FB4_RFID_Instance.Direccion_lectura;
   #Resultado := "FC_UDP_Bloque"(Id := 161, Origen := #Copia_161, Inicio := #Total, Foto := #Foto, Escritos := #Bloques_escritos, Final => #Total);
   #Copia_162 := "Est_DB_Gestor".FB4_RFID_Instance.Direccion_escritura;
   #Resultado := "FC_UDP_Bloque"(Id := 162, Origen := #Copia_162, Inicio := #Total, Foto := #Foto, Escritos := #Bloques_escritos, Final => #Total);
   #Copia_163 := "Est_DB_Gestor".FB4_RFID_Instance.Mascara_lectura;
   #Resultado := "FC_UDP_Bloque"(Id := 163, Origen := #Copia_163, Inicio := #Total, Foto := #Foto, Escritos := #Bloques_escritos, Final => #Total);
   #Copia_164 := "Est_DB_Gestor".FB4_RFID_Instance.Mascara_escritura;
   #Resultado := "FC_UDP_Bloque"(Id := 164, Origen := #Copia_164, Inicio := #Total, Foto := #Foto, Escritos := #Bloques_escritos, Final => #Total);
   #Copia_165 := "Est_DB_Gestor".FB4_RFID_Instance.Mascara_lectura_1;
   #Resultado := "FC_UDP_Bloque"(Id := 165, Origen := #Copia_165, Inicio := #Total, Foto := #Foto, Escritos := #Bloques_escritos, Final => #Total);
   #Copia_166 := "Est_DB_Gestor".FB4_RFID_Instance.Mascara_lectura_2;
   #Resultado := "FC_UDP_Bloque"(Id := 166, Origen := #Copia_166, Inicio := #Total, Foto := #Foto, Escritos := #Bloques_escritos, Final => #Total);
   #Copia_167 := "Est_DB_Gestor".FB4_RFID_Instance.Mascara_lectura_3;
   #Resultado := "FC_UDP_Bloque"(Id := 167, Origen := #Copia_167, Inicio := #Total, Foto := #Foto, Escritos := #Bloques_escritos, Final => #Total);
   #Copia_168 := "Est_DB_Gestor".FB4_RFID_Instance.Mascara_escritura_1;
   #Resultado := "FC_UDP_Bloque"(Id := 168, Origen := #Copia_168, Inicio := #Total, Foto := #Foto, Escritos := #Bloques_escritos, Final => #Total);
   #Copia_169 := "Est_DB_Gestor".FB4_RFID_Instance.Mascara_escritura_2;
   #Resultado := "FC_UDP_Bloque"(Id := 169, Origen := #Copia_169, Inicio := #Total, Foto := #Foto, Escritos := #Bloques_escritos, Final => #Total);
   #Copia_170 := "Est_DB_Gestor".FB4_RFID_Instance.Mascara_escritura_3;
   #Resultado := "FC_UDP_Bloque"(Id := 170, Origen := #Copia_170, Inicio := #Total, Foto := #Foto, Escritos := #Bloques_escritos, Final => #Total);
   #Copia_171 := "Est_DB_Gestor".FB4_RFID_Instance.T_Rfid.IN;
   #Resultado := "FC_UDP_Bloque"(Id := 171, Origen := #Copia_171, Inicio := #Total, Foto := #Foto, Escritos := #Bloques_escritos, Final => #Total);
   #Copia_172 := "Est_DB_Gestor".FB4_RFID_Instance.T_Rfid.Q;
   #Resultado := "FC_UDP_Bloque"(Id := 172, Origen := #Copia_172, Inicio := #Total, Foto := #Foto, Escritos := #Bloques_escritos, Final => #Total);
   #Copia_173 := "Est_DB_Gestor".FB4_RFID_Instance.T_Rfid.PT;
   #Resultado := "FC_UDP_Bloque"(Id := 173, Origen := #Copia_173, Inicio := #Total, Foto := #Foto, Escritos := #Bloques_escritos, Final => #Total);
   #Copia_174 := "Est_DB_Gestor".FB4_RFID_Instance.T_Rfid.ET;
   #Resultado := "FC_UDP_Bloque"(Id := 174, Origen := #Copia_174, Inicio := #Total, Foto := #Foto, Escritos := #Bloques_escritos, Final => #Total);
   #Copia_175 := "Est_DB_Gestor".FB4_RFID_Instance.Etapa_rfid;
   #Resultado := "FC_UDP_Bloque"(Id := 175, Origen := #Copia_175, Inicio := #Total, Foto := #Foto, Escritos := #Bloques_escritos, Final => #Total);
   #Copia_176 := "Est_DB_Gestor".FB4_RFID_Instance.Ventana_actual;
   #Resultado := "FC_UDP_Bloque"(Id := 176, Origen := #Copia_176, Inicio := #Total, Foto := #Foto, Escritos := #Bloques_escritos, Final => #Total);
   #Copia_177 := "Est_DB_Gestor".FB4_RFID_Instance.Mascara_lectura_tabla;
   #Resultado := "FC_UDP_Bloque"(Id := 177, Origen := #Copia_177, Inicio := #Total, Foto := #Foto, Escritos := #Bloques_escritos, Final => #Total);
   #Copia_178 := "Est_DB_Gestor".FB4_RFID_Instance.Mascara_escritura_tabla;
   #Resultado := "FC_UDP_Bloque"(Id := 178, Origen := #Copia_178, Inicio := #Total, Foto := #Foto, Escritos := #Bloques_escritos, Final => #Total);
   #Copia_179 := "Est_DB_Gestor".FB4_RFID_Instance.Ventana_lectura_activa;
   #Resultado := "FC_UDP_Bloque"(Id := 179, Origen := #Copia_179, Inicio := #Total, Foto := #Foto, Escritos := #Bloques_escritos, Final => #Total);
   #Copia_180 := "Est_DB_Gestor".FB4_RFID_Instance.Ventana_escritura_activa;
   #Resultado := "FC_UDP_Bloque"(Id := 180, Origen := #Copia_180, Inicio := #Total, Foto := #Foto, Escritos := #Bloques_escritos, Final => #Total);
   #Copia_181 := "Est_DB_Gestor".FB4_RFID_Instance.Direccion_ventana_lectura;
   #Resultado := "FC_UDP_Bloque"(Id := 181, Origen := #Copia_181, Inicio := #Total, Foto := #Foto, Escritos := #Bloques_escritos, Final => #Total);
   #Copia_182 := "Est_DB_Gestor".FB4_RFID_Instance.Direccion_ventana_escritura;
   #Resultado := "FC_UDP_Bloque"(Id := 182, Origen := #Copia_182, Inicio := #Total, Foto := #Foto, Escritos := #Bloques_escritos, Final => #Total);
   #Copia_183 := "Est_DB_Gestor".FB4_RFID_Instance.Etapa_7;
   #Resultado := "FC_UDP_Bloque"(Id := 183, Origen := #Copia_183, Inicio := #Total, Foto := #Foto, Escritos := #Bloques_escritos, Final => #Total);
   #Copia_184 := "Est_DB_Gestor".FB4_RFID_Instance.Etapa_9;
   #Resultado := "FC_UDP_Bloque"(Id := 184, Origen := #Copia_184, Inicio := #Total, Foto := #Foto, Escritos := #Bloques_escritos, Final => #Total);
   #Copia_185 := "Est_DB_Gestor".FB4_RFID_Instance.Etapa_1;
   #Resultado := "FC_UDP_Bloque"(Id := 185, Origen := #Copia_185, Inicio := #Total, Foto := #Foto, Escritos := #Bloques_escritos, Final => #Total);
   #Copia_186 := "Est_DB_Gestor".FB4_RFID_Instance.Etapa_3;
   #Resultado := "FC_UDP_Bloque"(Id := 186, Origen := #Copia_186, Inicio := #Total, Foto := #Foto, Escritos := #Bloques_escritos, Final => #Total);
   #Copia_187 := "Est_DB_Gestor".FB4_RFID_Instance.Etapa_4;
   #Resultado := "FC_UDP_Bloque"(Id := 187, Origen := #Copia_187, Inicio := #Total, Foto := #Foto, Escritos := #Bloques_escritos, Final => #Total);
   #Copia_188 := "Est_DB_Gestor".FB4_RFID_Instance.Rfid_ocupado;
   #Resultado := "FC_UDP_Bloque"(Id := 188, Origen := #Copia_188, Inicio := #Total, Foto := #Foto, Escritos := #Bloques_escritos, Final => #Total);
   #Copia_189 := "Est_DB_Gestor".FB4_RFID_Instance.Imagen_leida;
   #Resultado := "FC_UDP_Bloque"(Id := 189, Origen := #Copia_189, Inicio := #Total, Foto := #Foto, Escritos := #Bloques_escritos, Final => #Total);
   #Copia_190 := "Est_DB_Gestor".FB5_Reloj_Instance.Epoch_s;
   #Resultado := "FC_UDP_Bloque"(Id := 190, Origen := #Copia_190, Inicio := #Total, Foto := #Foto, Escritos := #Bloques_escritos, Final => #Total);
   #Copia_191 := "Est_DB_Gestor".FB5_Reloj_Instance.Milisegundos;
   #Resultado := "FC_UDP_Bloque"(Id := 191, Origen := #Copia_191, Inicio := #Total, Foto := #Foto, Escritos := #Bloques_escritos, Final => #Total);
   #Copia_192 := "Est_DB_Gestor".FB5_Reloj_Instance.Valida;
   #Resultado := "FC_UDP_Bloque"(Id := 192, Origen := #Copia_192, Inicio := #Total, Foto := #Foto, Escritos := #Bloques_escritos, Final => #Total);
   #Copia_193 := "Est_DB_Gestor".FB5_Reloj_Instance.Hora;
   #Resultado := "FC_UDP_Bloque"(Id := 193, Origen := #Copia_193, Inicio := #Total, Foto := #Foto, Escritos := #Bloques_escritos, Final => #Total);
   #Copia_194 := "Est_DB_Gestor".FB5_Reloj_Instance.Codigo;
   #Resultado := "FC_UDP_Bloque"(Id := 194, Origen := #Copia_194, Inicio := #Total, Foto := #Foto, Escritos := #Bloques_escritos, Final => #Total);
   #Copia_195 := "Est_DB_Gestor".FB5_Reloj_Instance.Anio;
   #Resultado := "FC_UDP_Bloque"(Id := 195, Origen := #Copia_195, Inicio := #Total, Foto := #Foto, Escritos := #Bloques_escritos, Final => #Total);
   #Copia_196 := "Est_DB_Gestor".FB5_Reloj_Instance.Mes;
   #Resultado := "FC_UDP_Bloque"(Id := 196, Origen := #Copia_196, Inicio := #Total, Foto := #Foto, Escritos := #Bloques_escritos, Final => #Total);
   #Copia_197 := "Est_DB_Gestor".FB5_Reloj_Instance.Dia;
   #Resultado := "FC_UDP_Bloque"(Id := 197, Origen := #Copia_197, Inicio := #Total, Foto := #Foto, Escritos := #Bloques_escritos, Final => #Total);
   #Copia_198 := "Est_DB_Gestor".FB5_Reloj_Instance.Era;
   #Resultado := "FC_UDP_Bloque"(Id := 198, Origen := #Copia_198, Inicio := #Total, Foto := #Foto, Escritos := #Bloques_escritos, Final => #Total);
   #Copia_199 := "Est_DB_Gestor".FB5_Reloj_Instance.Anio_era;
   #Resultado := "FC_UDP_Bloque"(Id := 199, Origen := #Copia_199, Inicio := #Total, Foto := #Foto, Escritos := #Bloques_escritos, Final => #Total);
   #Copia_200 := "Est_DB_Gestor".FB5_Reloj_Instance.Dia_anio;
   #Resultado := "FC_UDP_Bloque"(Id := 200, Origen := #Copia_200, Inicio := #Total, Foto := #Foto, Escritos := #Bloques_escritos, Final => #Total);
   #Copia_201 := "Est_DB_Gestor".FB5_Reloj_Instance.Dias;
   #Resultado := "FC_UDP_Bloque"(Id := 201, Origen := #Copia_201, Inicio := #Total, Foto := #Foto, Escritos := #Bloques_escritos, Final => #Total);
   #Copia_202 := "Est_DB_Gestor".Flanco_emergencia.CLK;
   #Resultado := "FC_UDP_Bloque"(Id := 202, Origen := #Copia_202, Inicio := #Total, Foto := #Foto, Escritos := #Bloques_escritos, Final => #Total);
   #Copia_203 := "Est_DB_Gestor".Flanco_emergencia.Q;
   #Resultado := "FC_UDP_Bloque"(Id := 203, Origen := #Copia_203, Inicio := #Total, Foto := #Foto, Escritos := #Bloques_escritos, Final => #Total);
   #Copia_204 := "Est_DB_Gestor".Etapa_gestion_anterior;
   #Resultado := "FC_UDP_Bloque"(Id := 204, Origen := #Copia_204, Inicio := #Total, Foto := #Foto, Escritos := #Bloques_escritos, Final => #Total);
   #Copia_205 := "Est_DB_Gestor".Emergencias_pendientes;
   #Resultado := "FC_UDP_Bloque"(Id := 205, Origen := #Copia_205, Inicio := #Total, Foto := #Foto, Escritos := #Bloques_escritos, Final => #Total);
   #Copia_206 := "Est_DB_Gestor".Inicio_app_segundos;
   #Resultado := "FC_UDP_Bloque"(Id := 206, Origen := #Copia_206, Inicio := #Total, Foto := #Foto, Escritos := #Bloques_escritos, Final => #Total);
   #Copia_207 := "Est_DB_Gestor".Inicio_app_milisegundos;
   #Resultado := "FC_UDP_Bloque"(Id := 207, Origen := #Copia_207, Inicio := #Total, Foto := #Foto, Escritos := #Bloques_escritos, Final => #Total);
   #Copia_208 := "Est_DB_Gestor".Ultima_secuencia;
   #Resultado := "FC_UDP_Bloque"(Id := 208, Origen := #Copia_208, Inicio := #Total, Foto := #Foto, Escritos := #Bloques_escritos, Final => #Total);
   #Copia_209 := "Est_DB_Gestor".Ciclo_manual_acabado;
   #Resultado := "FC_UDP_Bloque"(Id := 209, Origen := #Copia_209, Inicio := #Total, Foto := #Foto, Escritos := #Bloques_escritos, Final => #Total);
   #Copia_210 := "Est_DB_Gestor".Timer_parpadeo.IN;
   #Resultado := "FC_UDP_Bloque"(Id := 210, Origen := #Copia_210, Inicio := #Total, Foto := #Foto, Escritos := #Bloques_escritos, Final => #Total);
   #Copia_211 := "Est_DB_Gestor".Timer_parpadeo.Q;
   #Resultado := "FC_UDP_Bloque"(Id := 211, Origen := #Copia_211, Inicio := #Total, Foto := #Foto, Escritos := #Bloques_escritos, Final => #Total);
   #Copia_212 := "Est_DB_Gestor".Timer_parpadeo.PT;
   #Resultado := "FC_UDP_Bloque"(Id := 212, Origen := #Copia_212, Inicio := #Total, Foto := #Foto, Escritos := #Bloques_escritos, Final => #Total);
   #Copia_213 := "Est_DB_Gestor".Timer_parpadeo.ET;
   #Resultado := "FC_UDP_Bloque"(Id := 213, Origen := #Copia_213, Inicio := #Total, Foto := #Foto, Escritos := #Bloques_escritos, Final => #Total);
   #Copia_214 := "Est_DB_Gestor".Parpadeo;
   #Resultado := "FC_UDP_Bloque"(Id := 214, Origen := #Copia_214, Inicio := #Total, Foto := #Foto, Escritos := #Bloques_escritos, Final => #Total);
   #Copia_215 := "FB_App_Camara_DB".App_inicio;
   #Resultado := "FC_UDP_Bloque"(Id := 215, Origen := #Copia_215, Inicio := #Total, Foto := #Foto, Escritos := #Bloques_escritos, Final => #Total);
   #Copia_216 := "FB_App_Camara_DB".Emergencia;
   #Resultado := "FC_UDP_Bloque"(Id := 216, Origen := #Copia_216, Inicio := #Total, Foto := #Foto, Escritos := #Bloques_escritos, Final => #Total);
   #Copia_217 := "FB_App_Camara_DB".Estado_camara;
   #Resultado := "FC_UDP_Bloque"(Id := 217, Origen := #Copia_217, Inicio := #Total, Foto := #Foto, Escritos := #Bloques_escritos, Final => #Total);
   #Copia_218 := "FB_App_Camara_DB".Entradas_camara;
   #Resultado := "FC_UDP_Bloque"(Id := 218, Origen := #Copia_218, Inicio := #Total, Foto := #Foto, Escritos := #Bloques_escritos, Final => #Total);
   #Copia_219 := "FB_App_Camara_DB".App_en_reposo;
   #Resultado := "FC_UDP_Bloque"(Id := 219, Origen := #Copia_219, Inicio := #Total, Foto := #Foto, Escritos := #Bloques_escritos, Final => #Total);
   #Copia_220 := "FB_App_Camara_DB".App_terminada;
   #Resultado := "FC_UDP_Bloque"(Id := 220, Origen := #Copia_220, Inicio := #Total, Foto := #Foto, Escritos := #Bloques_escritos, Final => #Total);
   #Copia_221 := "FB_App_Camara_DB".App_alarma;
   #Resultado := "FC_UDP_Bloque"(Id := 221, Origen := #Copia_221, Inicio := #Total, Foto := #Foto, Escritos := #Bloques_escritos, Final => #Total);
   #Copia_222 := "FB_App_Camara_DB".App_rearme_requerido;
   #Resultado := "FC_UDP_Bloque"(Id := 222, Origen := #Copia_222, Inicio := #Total, Foto := #Foto, Escritos := #Bloques_escritos, Final => #Total);
   #Copia_223 := "FB_App_Camara_DB".Inhibir_cinta;
   #Resultado := "FC_UDP_Bloque"(Id := 223, Origen := #Copia_223, Inicio := #Total, Foto := #Foto, Escritos := #Bloques_escritos, Final => #Total);
   #Copia_224 := "FB_App_Camara_DB".Mando_camara;
   #Resultado := "FC_UDP_Bloque"(Id := 224, Origen := #Copia_224, Inicio := #Total, Foto := #Foto, Escritos := #Bloques_escritos, Final => #Total);
   #Copia_225 := "FB_App_Camara_DB".Salidas_camara;
   #Resultado := "FC_UDP_Bloque"(Id := 225, Origen := #Copia_225, Inicio := #Total, Foto := #Foto, Escritos := #Bloques_escritos, Final => #Total);
   #Copia_226 := "FB_App_Camara_DB".Etapa_app;
   #Resultado := "FC_UDP_Bloque"(Id := 226, Origen := #Copia_226, Inicio := #Total, Foto := #Foto, Escritos := #Bloques_escritos, Final => #Total);
   #Copia_227 := "FB_App_Camara_DB".Job_actual;
   #Resultado := "FC_UDP_Bloque"(Id := 227, Origen := #Copia_227, Inicio := #Total, Foto := #Foto, Escritos := #Bloques_escritos, Final => #Total);
   #Copia_228 := "FB_App_Camara_DB".Orden_a_run;
   #Resultado := "FC_UDP_Bloque"(Id := 228, Origen := #Copia_228, Inicio := #Total, Foto := #Foto, Escritos := #Bloques_escritos, Final => #Total);
   #Copia_229 := "FB_App_Camara_DB".Orden_cambio_job;
   #Resultado := "FC_UDP_Bloque"(Id := 229, Origen := #Copia_229, Inicio := #Total, Foto := #Foto, Escritos := #Bloques_escritos, Final => #Total);
   #Copia_230 := "FB_App_Camara_DB".Orden_disparo;
   #Resultado := "FC_UDP_Bloque"(Id := 230, Origen := #Copia_230, Inicio := #Total, Foto := #Foto, Escritos := #Bloques_escritos, Final => #Total);
   #Copia_231 := "FB_App_Camara_DB".Fallo_camara;
   #Resultado := "FC_UDP_Bloque"(Id := 231, Origen := #Copia_231, Inicio := #Total, Foto := #Foto, Escritos := #Bloques_escritos, Final => #Total);
   #Copia_232 := "FB_App_Camara_DB".Flanco_ack_run.CLK;
   #Resultado := "FC_UDP_Bloque"(Id := 232, Origen := #Copia_232, Inicio := #Total, Foto := #Foto, Escritos := #Bloques_escritos, Final => #Total);
   #Copia_233 := "FB_App_Camara_DB".Flanco_ack_run.Q;
   #Resultado := "FC_UDP_Bloque"(Id := 233, Origen := #Copia_233, Inicio := #Total, Foto := #Foto, Escritos := #Bloques_escritos, Final => #Total);
   #Copia_234 := "FB_App_Camara_DB".Flanco_ack_job.CLK;
   #Resultado := "FC_UDP_Bloque"(Id := 234, Origen := #Copia_234, Inicio := #Total, Foto := #Foto, Escritos := #Bloques_escritos, Final => #Total);
   #Copia_235 := "FB_App_Camara_DB".Flanco_ack_job.Q;
   #Resultado := "FC_UDP_Bloque"(Id := 235, Origen := #Copia_235, Inicio := #Total, Foto := #Foto, Escritos := #Bloques_escritos, Final => #Total);
   #Copia_236 := "FB_App_Camara_DB".Flanco_ready.CLK;
   #Resultado := "FC_UDP_Bloque"(Id := 236, Origen := #Copia_236, Inicio := #Total, Foto := #Foto, Escritos := #Bloques_escritos, Final => #Total);
   #Copia_237 := "FB_App_Camara_DB".Flanco_ready.Q;
   #Resultado := "FC_UDP_Bloque"(Id := 237, Origen := #Copia_237, Inicio := #Total, Foto := #Foto, Escritos := #Bloques_escritos, Final => #Total);
   #Copia_238 := "FB_App_Camara_DB".Pulso_a_run.IN;
   #Resultado := "FC_UDP_Bloque"(Id := 238, Origen := #Copia_238, Inicio := #Total, Foto := #Foto, Escritos := #Bloques_escritos, Final => #Total);
   #Copia_239 := "FB_App_Camara_DB".Pulso_a_run.Q;
   #Resultado := "FC_UDP_Bloque"(Id := 239, Origen := #Copia_239, Inicio := #Total, Foto := #Foto, Escritos := #Bloques_escritos, Final => #Total);
   #Copia_240 := "FB_App_Camara_DB".Pulso_a_run.PT;
   #Resultado := "FC_UDP_Bloque"(Id := 240, Origen := #Copia_240, Inicio := #Total, Foto := #Foto, Escritos := #Bloques_escritos, Final => #Total);
   #Copia_241 := "FB_App_Camara_DB".Pulso_a_run.ET;
   #Resultado := "FC_UDP_Bloque"(Id := 241, Origen := #Copia_241, Inicio := #Total, Foto := #Foto, Escritos := #Bloques_escritos, Final => #Total);
   #Copia_242 := "FB_App_Camara_DB".Pulso_cambio_job.IN;
   #Resultado := "FC_UDP_Bloque"(Id := 242, Origen := #Copia_242, Inicio := #Total, Foto := #Foto, Escritos := #Bloques_escritos, Final => #Total);
   #Copia_243 := "FB_App_Camara_DB".Pulso_cambio_job.Q;
   #Resultado := "FC_UDP_Bloque"(Id := 243, Origen := #Copia_243, Inicio := #Total, Foto := #Foto, Escritos := #Bloques_escritos, Final => #Total);
   #Copia_244 := "FB_App_Camara_DB".Pulso_cambio_job.PT;
   #Resultado := "FC_UDP_Bloque"(Id := 244, Origen := #Copia_244, Inicio := #Total, Foto := #Foto, Escritos := #Bloques_escritos, Final => #Total);
   #Copia_245 := "FB_App_Camara_DB".Pulso_cambio_job.ET;
   #Resultado := "FC_UDP_Bloque"(Id := 245, Origen := #Copia_245, Inicio := #Total, Foto := #Foto, Escritos := #Bloques_escritos, Final => #Total);
   #Copia_246 := "FB_App_Camara_DB".Pulso_disparo.IN;
   #Resultado := "FC_UDP_Bloque"(Id := 246, Origen := #Copia_246, Inicio := #Total, Foto := #Foto, Escritos := #Bloques_escritos, Final => #Total);
   #Copia_247 := "FB_App_Camara_DB".Pulso_disparo.Q;
   #Resultado := "FC_UDP_Bloque"(Id := 247, Origen := #Copia_247, Inicio := #Total, Foto := #Foto, Escritos := #Bloques_escritos, Final => #Total);
   #Copia_248 := "FB_App_Camara_DB".Pulso_disparo.PT;
   #Resultado := "FC_UDP_Bloque"(Id := 248, Origen := #Copia_248, Inicio := #Total, Foto := #Foto, Escritos := #Bloques_escritos, Final => #Total);
   #Copia_249 := "FB_App_Camara_DB".Pulso_disparo.ET;
   #Resultado := "FC_UDP_Bloque"(Id := 249, Origen := #Copia_249, Inicio := #Total, Foto := #Foto, Escritos := #Bloques_escritos, Final => #Total);
   #Copia_250 := "FB_App_Camara_DB".Temporizador_camara.IN;
   #Resultado := "FC_UDP_Bloque"(Id := 250, Origen := #Copia_250, Inicio := #Total, Foto := #Foto, Escritos := #Bloques_escritos, Final => #Total);
   #Copia_251 := "FB_App_Camara_DB".Temporizador_camara.Q;
   #Resultado := "FC_UDP_Bloque"(Id := 251, Origen := #Copia_251, Inicio := #Total, Foto := #Foto, Escritos := #Bloques_escritos, Final => #Total);
   #Copia_252 := "FB_App_Camara_DB".Temporizador_camara.PT;
   #Resultado := "FC_UDP_Bloque"(Id := 252, Origen := #Copia_252, Inicio := #Total, Foto := #Foto, Escritos := #Bloques_escritos, Final => #Total);
   #Copia_253 := "FB_App_Camara_DB".Temporizador_camara.ET;
   #Resultado := "FC_UDP_Bloque"(Id := 253, Origen := #Copia_253, Inicio := #Total, Foto := #Foto, Escritos := #Bloques_escritos, Final => #Total);
   #Copia_254 := "FB_App_Camara_DB".Temporizador_verde.IN;
   #Resultado := "FC_UDP_Bloque"(Id := 254, Origen := #Copia_254, Inicio := #Total, Foto := #Foto, Escritos := #Bloques_escritos, Final => #Total);
   #Copia_255 := "FB_App_Camara_DB".Temporizador_verde.Q;
   #Resultado := "FC_UDP_Bloque"(Id := 255, Origen := #Copia_255, Inicio := #Total, Foto := #Foto, Escritos := #Bloques_escritos, Final => #Total);
   #Copia_256 := "FB_App_Camara_DB".Temporizador_verde.PT;
   #Resultado := "FC_UDP_Bloque"(Id := 256, Origen := #Copia_256, Inicio := #Total, Foto := #Foto, Escritos := #Bloques_escritos, Final => #Total);
   #Copia_257 := "FB_App_Camara_DB".Temporizador_verde.ET;
   #Resultado := "FC_UDP_Bloque"(Id := 257, Origen := #Copia_257, Inicio := #Total, Foto := #Foto, Escritos := #Bloques_escritos, Final => #Total);
   #Copia_258 := "FB_App_Camara_DB".Temporizador_rojo.IN;
   #Resultado := "FC_UDP_Bloque"(Id := 258, Origen := #Copia_258, Inicio := #Total, Foto := #Foto, Escritos := #Bloques_escritos, Final => #Total);
   #Copia_259 := "FB_App_Camara_DB".Temporizador_rojo.Q;
   #Resultado := "FC_UDP_Bloque"(Id := 259, Origen := #Copia_259, Inicio := #Total, Foto := #Foto, Escritos := #Bloques_escritos, Final => #Total);
   #Copia_260 := "FB_App_Camara_DB".Temporizador_rojo.PT;
   #Resultado := "FC_UDP_Bloque"(Id := 260, Origen := #Copia_260, Inicio := #Total, Foto := #Foto, Escritos := #Bloques_escritos, Final => #Total);
   #Copia_261 := "FB_App_Camara_DB".Temporizador_rojo.ET;
   #Resultado := "FC_UDP_Bloque"(Id := 261, Origen := #Copia_261, Inicio := #Total, Foto := #Foto, Escritos := #Bloques_escritos, Final => #Total);
   #Copia_262 := "Profinet_ctrl";
   #Resultado := "FC_UDP_Bloque"(Id := 262, Origen := #Copia_262, Inicio := #Total, Foto := #Foto, Escritos := #Bloques_escritos, Final => #Total);
   #Copia_263 := "Profinet_status";
   #Resultado := "FC_UDP_Bloque"(Id := 263, Origen := #Copia_263, Inicio := #Total, Foto := #Foto, Escritos := #Bloques_escritos, Final => #Total);
   #Copia_264 := "Clock_Byte";
   #Resultado := "FC_UDP_Bloque"(Id := 264, Origen := #Copia_264, Inicio := #Total, Foto := #Foto, Escritos := #Bloques_escritos, Final => #Total);
   #Copia_265 := "Clock_10Hz";
   #Resultado := "FC_UDP_Bloque"(Id := 265, Origen := #Copia_265, Inicio := #Total, Foto := #Foto, Escritos := #Bloques_escritos, Final => #Total);
   #Copia_266 := "Clock_5Hz";
   #Resultado := "FC_UDP_Bloque"(Id := 266, Origen := #Copia_266, Inicio := #Total, Foto := #Foto, Escritos := #Bloques_escritos, Final => #Total);
   #Copia_267 := "Clock_2.5Hz";
   #Resultado := "FC_UDP_Bloque"(Id := 267, Origen := #Copia_267, Inicio := #Total, Foto := #Foto, Escritos := #Bloques_escritos, Final => #Total);
   #Copia_268 := "Clock_2Hz";
   #Resultado := "FC_UDP_Bloque"(Id := 268, Origen := #Copia_268, Inicio := #Total, Foto := #Foto, Escritos := #Bloques_escritos, Final => #Total);
   #Copia_269 := "Clock_1.25Hz";
   #Resultado := "FC_UDP_Bloque"(Id := 269, Origen := #Copia_269, Inicio := #Total, Foto := #Foto, Escritos := #Bloques_escritos, Final => #Total);
   #Copia_270 := "Clock_1Hz";
   #Resultado := "FC_UDP_Bloque"(Id := 270, Origen := #Copia_270, Inicio := #Total, Foto := #Foto, Escritos := #Bloques_escritos, Final => #Total);
   #Copia_271 := "Clock_0.625Hz";
   #Resultado := "FC_UDP_Bloque"(Id := 271, Origen := #Copia_271, Inicio := #Total, Foto := #Foto, Escritos := #Bloques_escritos, Final => #Total);
   #Copia_272 := "Clock_0.5Hz";
   #Resultado := "FC_UDP_Bloque"(Id := 272, Origen := #Copia_272, Inicio := #Total, Foto := #Foto, Escritos := #Bloques_escritos, Final => #Total);
   #Copia_273 := "Entradas_APP";
   #Resultado := "FC_UDP_Bloque"(Id := 273, Origen := #Copia_273, Inicio := #Total, Foto := #Foto, Escritos := #Bloques_escritos, Final => #Total);
   #Copia_274 := "Entradas_Basico";
   #Resultado := "FC_UDP_Bloque"(Id := 274, Origen := #Copia_274, Inicio := #Total, Foto := #Foto, Escritos := #Bloques_escritos, Final => #Total);
   #Copia_275 := "Entradas_Stopper";
   #Resultado := "FC_UDP_Bloque"(Id := 275, Origen := #Copia_275, Inicio := #Total, Foto := #Foto, Escritos := #Bloques_escritos, Final => #Total);
   #Copia_276 := "Salidas_Basico";
   #Resultado := "FC_UDP_Bloque"(Id := 276, Origen := #Copia_276, Inicio := #Total, Foto := #Foto, Escritos := #Bloques_escritos, Final => #Total);
   #Copia_277 := "Salidas_APP";
   #Resultado := "FC_UDP_Bloque"(Id := 277, Origen := #Copia_277, Inicio := #Total, Foto := #Foto, Escritos := #Bloques_escritos, Final => #Total);
   #Copia_278 := "Entradas_RFID";
   #Resultado := "FC_UDP_Bloque"(Id := 278, Origen := #Copia_278, Inicio := #Total, Foto := #Foto, Escritos := #Bloques_escritos, Final => #Total);
   #Copia_279 := "Salidas_RFID";
   #Resultado := "FC_UDP_Bloque"(Id := 279, Origen := #Copia_279, Inicio := #Total, Foto := #Foto, Escritos := #Bloques_escritos, Final => #Total);
   #Bloques_omitidos := #N_BLOQUES - #Bloques_escritos;
   #Cursor := 0;
   #Etapa := 2;
END_IF;

// un datagrama por trozo: cabecera de 18 bytes + bloques enteros (id, longitud, datos)
IF #Etapa = 2 THEN
   #Bytes_trozo := 0;
   #Bloques_trozo := 0;
   #longitud := #Cursor;
   WHILE #Cursor < #Total DO
      #lon_bloque := BYTE_TO_DINT(#Foto[#Cursor + 2]) * 256 + BYTE_TO_DINT(#Foto[#Cursor + 3]) + 4;
      IF #Bytes_trozo + #lon_bloque > #MAX_PAYLOAD AND #Bloques_trozo > 0 THEN EXIT; END_IF;
      #Bytes_trozo := #Bytes_trozo + #lon_bloque;
      #Cursor := #Cursor + #lon_bloque;
      #Bloques_trozo := #Bloques_trozo + 1;
   END_WHILE;
   #Datagrama[0] := 16#50;
   #Datagrama[1] := 16#47;
   #Datagrama[2] := 2;
   #Datagrama[3] := USINT_TO_BYTE(#ID_PLC);
   #d := UDINT_TO_DWORD(#Secuencia);
   #Datagrama[4] := #d.%B3;
   #Datagrama[5] := #d.%B2;
   #Datagrama[6] := #d.%B1;
   #Datagrama[7] := #d.%B0;
   #l := LINT_TO_LWORD(#Marca_tiempo);
   #Datagrama[8] := #l.%B7;
   #Datagrama[9] := #l.%B6;
   #Datagrama[10] := #l.%B5;
   #Datagrama[11] := #l.%B4;
   #Datagrama[12] := #l.%B3;
   #Datagrama[13] := #l.%B2;
   #Datagrama[14] := #l.%B1;
   #Datagrama[15] := #l.%B0;
   #w := UINT_TO_WORD(#Bloques_trozo);
   #Datagrama[16] := #w.%B1;
   #Datagrama[17] := #w.%B0;
   #resultado := MOVE_BLK_VARIANT(SRC := #Foto, COUNT := DINT_TO_UDINT(#Bytes_trozo),
                                  SRC_INDEX := #longitud, DEST_INDEX := 18, DEST => #Datagrama);
   #Secuencia := #Secuencia + 1;
   #Lanza_envio := TRUE;
   #Etapa := 3;
END_IF;

#Cliente_envio(REQ := #Lanza_envio, ID := #Conexion.ID, LEN := DINT_TO_UDINT(#Bytes_trozo + 18),
               DATA := #Datagrama, ADDR := #Destino, STATUS => #Estado_tusend);
#Lanza_envio := FALSE;

// resultado del envio; si la conexion se perdio, a reconectar
#Espera_envio(IN := #Etapa = 3, PT := T#1s);
IF #Etapa = 3 THEN
   IF #Cliente_envio.DONE THEN
      #Enviados := #Enviados + 1;
      IF #Cursor >= #Total THEN #Etapa := 1; ELSE #Etapa := 2; END_IF;
   ELSIF #Cliente_envio.ERROR OR #Espera_envio.Q THEN
      #Fallidos := #Fallidos + 1;
      #Conectado := FALSE;
      #Etapa := 0;
   END_IF;
END_IF;

END_FUNCTION_BLOCK
